// Tests for MONETcommon.FB_MonetTempSensor, the scaling and wire-break check of the 0-10 V temperature sensors.
// Cabinet_Over_Temp_Requests_Roof_Close: the cabinet temperature thresholds of MONETcommon.FB_MonetCabinetControl (BT1, driven
// through FB_MonetCabinetProbe) and its bCloseRoofRequest (#24 D9); no telescope is passed, so nothing is parked.
// Cabinet_Reads_The_Key_And_Passes_The_Safety_Inputs: FB_MonetCabinetControl as BROTLib.I_Cabinet (X1).
// Safety_Items_Decode_The_Info_Blocks: FB_MonetSafetyHandling as BROTLib.I_SafetyDiagnostics (X4), driven through FB_MonetSafetyProbe.
FUNCTION_BLOCK FB_MonetTempSensor_Tests EXTENDS TcUnit.FB_TestSuite
VAR
	nullComm	: FB_NullComm;
END_VAR

Mid_Scale_Is_Valid();
Wire_Break_Is_Invalid();
Over_Range_Is_Invalid();
Recovers_After_Wire_Break();
Cabinet_Over_Temp_Requests_Roof_Close();
Cabinet_Reads_The_Key_And_Passes_The_Safety_Inputs();
Safety_Items_Decode_The_Info_Blocks();

// 16384 of 32767 is 5 V, i.e. 25 C.
METHOD PRIVATE Mid_Scale_Is_Valid
VAR
	sensor	: MONETcommon.FB_MonetTempSensor;
END_VAR
TEST('Mid_Scale_Is_Valid');
sensor(iRaw := 16384, sName := 'TEMP_M1', comm := nullComm);
AssertTrue(Condition := sensor.bValid, Message := 'valid');
AssertEquals_REAL(Expected := 25.0, Actual := sensor.fTemperature, Delta := 0.01, Message := 'temperature');
TEST_FINISHED();
END_METHOD

// A broken wire reads about 0 V, which scales to -50 C.
METHOD PRIVATE Wire_Break_Is_Invalid
VAR
	sensor	: MONETcommon.FB_MonetTempSensor;
END_VAR
TEST('Wire_Break_Is_Invalid');
sensor(iRaw := 0, sName := 'TEMP_M1', comm := nullComm);
AssertFalse(Condition := sensor.bValid, Message := 'raw 0');
sensor(iRaw := 327, sName := 'TEMP_M1', comm := nullComm);
AssertFalse(Condition := sensor.bValid, Message := 'raw 327, just below 1 %');
sensor(iRaw := 328, sName := 'TEMP_M1', comm := nullComm);
AssertTrue(Condition := sensor.bValid, Message := 'raw 328, 1 %');
TEST_FINISHED();
END_METHOD

METHOD PRIVATE Over_Range_Is_Invalid
VAR
	sensor	: MONETcommon.FB_MonetTempSensor;
END_VAR
TEST('Over_Range_Is_Invalid');
sensor(iRaw := 32766, sName := 'TEMP_M1', comm := nullComm);
AssertTrue(Condition := sensor.bValid, Message := 'raw 32766');
sensor(iRaw := 32767, sName := 'TEMP_M1', comm := nullComm);
AssertFalse(Condition := sensor.bValid, Message := 'raw 32767, full scale');
TEST_FINISHED();
END_METHOD

METHOD PRIVATE Recovers_After_Wire_Break
VAR
	sensor	: MONETcommon.FB_MonetTempSensor;
END_VAR
TEST('Recovers_After_Wire_Break');
sensor(iRaw := 0, sName := 'TEMP_M1', comm := nullComm);
AssertFalse(Condition := sensor.bValid, Message := 'broken');
sensor(iRaw := 16384, sName := 'TEMP_M1', comm := nullComm);
AssertTrue(Condition := sensor.bValid, Message := 'reconnected');
TEST_FINISHED();
END_METHOD

// #24 D9 (owner decision: a critical cabinet temperature parks everything, the roof included): bCloseRoofRequest equals
// bCabinetOverTemp, set above 60 C and held until below 50 C, not latched beyond that. One call per temperature (BT1 in
// 0.1 C), no telescope (iTelescope 0).
METHOD PRIVATE Cabinet_Over_Temp_Requests_Roof_Close
VAR
	fbComm	: FB_NullComm;
	fbCab	: FB_MonetCabinetProbe(comm := fbComm);
END_VAR
TEST('Cabinet_Over_Temp_Requests_Roof_Close');
fbCab(fCabinetTempIn := 25.0);
AssertFalse(Condition := fbCab.bCloseRoofRequest, Message := '25 C: no roof close request');
fbCab(fCabinetTempIn := 59.9);
AssertFalse(Condition := fbCab.bCloseRoofRequest, Message := '59.9 C on the way up: no roof close request');
AssertFalse(Condition := fbCab.bCabinetOverTemp, Message := '59.9 C on the way up: not over temperature');
fbCab(fCabinetTempIn := 60.1);
AssertTrue(Condition := fbCab.bCloseRoofRequest, Message := '60.1 C: roof close requested');
AssertTrue(Condition := fbCab.bCabinetOverTemp, Message := '60.1 C: over temperature');
fbCab(fCabinetTempIn := 55.0);
AssertTrue(Condition := fbCab.bCloseRoofRequest, Message := '55 C on the way down: the request holds');
fbCab(fCabinetTempIn := 50.0);
AssertTrue(Condition := fbCab.bCloseRoofRequest, Message := '50.0 C on the way down: the request holds (reset below 50)');
fbCab(fCabinetTempIn := 49.9);
AssertFalse(Condition := fbCab.bCloseRoofRequest, Message := '49.9 C: the request is gone');
AssertFalse(Condition := fbCab.bCabinetOverTemp, Message := '49.9 C: not over temperature');
fbCab(fCabinetTempIn := 55.0);
AssertFalse(Condition := fbCab.bCloseRoofRequest, Message := '55 C on the way up again: no latch, no request');
TEST_FINISHED();
END_METHOD

// X1: ControlMode follows the Local/Remote key (inKeyLocal TRUE = Local), SwitchPresent is TRUE, the four other properties are the inputs.
METHOD PRIVATE Cabinet_Reads_The_Key_And_Passes_The_Safety_Inputs
VAR
	fbComm	: FB_NullComm;
	fbCab	: FB_MonetCabinetProbe(comm := fbComm);
	ipCab	: BROTLib.I_Cabinet;
END_VAR
TEST('Cabinet_Reads_The_Key_And_Passes_The_Safety_Inputs');
ipCab := fbCab;
fbCab(fCabinetTempIn := 25.0, bKeyLocalIn := FALSE, bEstop := FALSE, bSafetyError := FALSE, bSafetyAckPending := FALSE, bPendantActive := FALSE);
AssertTrue(Condition := ipCab.ControlMode = BROTLib.E_ControlMode.remote, Message := 'key off: Remote');
AssertTrue(Condition := ipCab.SwitchPresent, Message := 'the key is a physical switch');
AssertFalse(Condition := ipCab.EstopActive OR ipCab.SafetyError OR ipCab.SafetyAckPending OR ipCab.PendantActive, Message := 'inputs at rest: all FALSE');
fbCab(fCabinetTempIn := 25.0, bKeyLocalIn := TRUE, bEstop := FALSE, bSafetyError := FALSE, bSafetyAckPending := FALSE, bPendantActive := FALSE);
AssertTrue(Condition := ipCab.ControlMode = BROTLib.E_ControlMode.local, Message := 'key on: Local');
fbCab(fCabinetTempIn := 25.0, bKeyLocalIn := FALSE, bEstop := TRUE, bSafetyError := FALSE, bSafetyAckPending := FALSE, bPendantActive := FALSE);
AssertTrue(Condition := ipCab.EstopActive AND NOT ipCab.SafetyError AND NOT ipCab.SafetyAckPending AND NOT ipCab.PendantActive, Message := 'only EstopActive');
fbCab(fCabinetTempIn := 25.0, bKeyLocalIn := FALSE, bEstop := FALSE, bSafetyError := TRUE, bSafetyAckPending := FALSE, bPendantActive := FALSE);
AssertTrue(Condition := ipCab.SafetyError AND NOT ipCab.EstopActive AND NOT ipCab.SafetyAckPending AND NOT ipCab.PendantActive, Message := 'only SafetyError');
fbCab(fCabinetTempIn := 25.0, bKeyLocalIn := FALSE, bEstop := FALSE, bSafetyError := FALSE, bSafetyAckPending := TRUE, bPendantActive := FALSE);
AssertTrue(Condition := ipCab.SafetyAckPending AND NOT ipCab.EstopActive AND NOT ipCab.SafetyError AND NOT ipCab.PendantActive, Message := 'only SafetyAckPending');
fbCab(fCabinetTempIn := 25.0, bKeyLocalIn := FALSE, bEstop := FALSE, bSafetyError := FALSE, bSafetyAckPending := FALSE, bPendantActive := TRUE);
AssertTrue(Condition := ipCab.PendantActive AND NOT ipCab.EstopActive AND NOT ipCab.SafetyError AND NOT ipCab.SafetyAckPending, Message := 'only PendantActive');
TEST_FINISHED();
END_METHOD

// X4: items, texts, raw bytes, bOk, RestartPending (state RESET) and the derived StoActive, through the info data of the TwinSAFE blocks.
METHOD PRIVATE Safety_Items_Decode_The_Info_Blocks
VAR
	fbComm	: FB_NullComm;
	fbSafe	: FB_MonetSafetyProbe(comm := fbComm);
	ipSafe	: BROTLib.I_SafetyDiagnostics;
	stItems	: BROTLib.ST_SafetyItems;
END_VAR
TEST('Safety_Items_Decode_The_Info_Blocks');
ipSafe := fbSafe;
// everything in its normal running state
fbSafe(nGroupState := 1, nEStopState := 1, nEStopDiag := 0, nInState := 104, nInDiag := 0, nInSignals := 0, nOutState := 104, nOutDiag := 0, nOutSignals := 0);
stItems := ipSafe.Items;
AssertTrue(Condition := stItems.nCount = 4, Message := 'four items');
AssertEquals_STRING(Expected := 'safety.group1', Actual := stItems.aItem[1].sName, Message := 'item 1 name');
AssertEquals_STRING(Expected := 'safety.estop1', Actual := stItems.aItem[2].sName, Message := 'item 2 name');
AssertEquals_STRING(Expected := 'safety.el1904', Actual := stItems.aItem[3].sName, Message := 'item 3 name');
AssertEquals_STRING(Expected := 'safety.el2904', Actual := stItems.aItem[4].sName, Message := 'item 4 name');
AssertTrue(Condition := stItems.aItem[1].eKind = BROTLib.E_SafetyItemKind.group AND stItems.aItem[2].eKind = BROTLib.E_SafetyItemKind.estop
	AND stItems.aItem[3].eKind = BROTLib.E_SafetyItemKind.connection_in AND stItems.aItem[4].eKind = BROTLib.E_SafetyItemKind.connection_out, Message := 'kinds');
AssertTrue(Condition := stItems.aItem[1].bOk AND stItems.aItem[2].bOk AND stItems.aItem[3].bOk AND stItems.aItem[4].bOk, Message := 'all ok in the normal state');
AssertEquals_STRING(Expected := 'RUN', Actual := stItems.aItem[1].sState, Message := 'group state text');
AssertEquals_STRING(Expected := 'State Data', Actual := stItems.aItem[3].sState, Message := 'connection state text');
AssertFalse(Condition := ipSafe.StoActive, Message := 'no STO in the normal state');
AssertFalse(Condition := ipSafe.RestartPending, Message := 'no restart pending in the normal state');
// E-stop pressed: state STOP
fbSafe(nGroupState := 1, nEStopState := 2, nEStopDiag := 0, nInState := 104, nInDiag := 0, nInSignals := 0, nOutState := 104, nOutDiag := 0, nOutSignals := 0);
stItems := ipSafe.Items;
AssertFalse(Condition := stItems.aItem[2].bOk, Message := 'E-stop item not ok');
AssertEquals_STRING(Expected := 'STOP', Actual := stItems.aItem[2].sState, Message := 'E-stop state text');
AssertTrue(Condition := stItems.aItem[2].nMapState = 2, Message := 'raw E-stop map state');
AssertTrue(Condition := stItems.aItem[1].bOk, Message := 'the group item is not affected');
AssertTrue(Condition := ipSafe.StoActive, Message := 'STO derived from the E-stop not in RUN');
AssertFalse(Condition := ipSafe.RestartPending, Message := 'STOP is not RESET');
// group waits for restart: state RESET (also with the E-stop function)
fbSafe(nGroupState := 5, nEStopState := 5, nEStopDiag := 0, nInState := 104, nInDiag := 0, nInSignals := 0, nOutState := 104, nOutDiag := 0, nOutSignals := 0);
stItems := ipSafe.Items;
AssertTrue(Condition := ipSafe.RestartPending, Message := 'RESET: restart pending');
AssertEquals_STRING(Expected := 'RESET', Actual := stItems.aItem[1].sState, Message := 'group state text RESET');
AssertFalse(Condition := stItems.aItem[1].bOk, Message := 'group item not ok in RESET');
AssertTrue(Condition := ipSafe.StoActive, Message := 'STO derived');
// only the E-stop function waits
fbSafe(nGroupState := 1, nEStopState := 5, nEStopDiag := 0, nInState := 104, nInDiag := 0, nInSignals := 0, nOutState := 104, nOutDiag := 0, nOutSignals := 0);
AssertTrue(Condition := ipSafe.RestartPending, Message := 'E-stop RESET alone: restart pending');
// a diagnosis on the E-stop makes it not ok even in RUN
fbSafe(nGroupState := 1, nEStopState := 1, nEStopDiag := 16, nInState := 104, nInDiag := 0, nInSignals := 0, nOutState := 104, nOutDiag := 0, nOutSignals := 0);
stItems := ipSafe.Items;
AssertFalse(Condition := stItems.aItem[2].bOk, Message := 'E-stop diagnosis: not ok');
AssertEquals_STRING(Expected := 'EDM Error EDM 1', Actual := stItems.aItem[2].sDiag, Message := 'E-stop diagnosis text');
// connections: diagnosis, channel bits (low nibble only), other state
fbSafe(nGroupState := 1, nEStopState := 1, nEStopDiag := 0, nInState := 104, nInDiag := 5, nInSignals := 245, nOutState := 103, nOutDiag := 0, nOutSignals := 0);
stItems := ipSafe.Items;
AssertFalse(Condition := stItems.aItem[3].bOk, Message := 'EL1904 diagnosis: not ok');
AssertEquals_STRING(Expected := 'Watchdog expired', Actual := stItems.aItem[3].sDiag, Message := 'EL1904 diagnosis text');
AssertTrue(Condition := stItems.aItem[3].nChannels = 16#05, Message := 'EL1904 channels 1 and 3');
AssertTrue(Condition := stItems.aItem[3].nMapDiag = 16#05, Message := 'raw EL1904 diagnosis');
AssertFalse(Condition := stItems.aItem[4].bOk, Message := 'EL2904 not in State Data');
AssertEquals_STRING(Expected := 'State Parameter', Actual := stItems.aItem[4].sState, Message := 'EL2904 state text');
TEST_FINISHED();
END_METHOD

END_FUNCTION_BLOCK

(* stored: Version 1.1.0.1, ProductVersion 3.1.4024.15
   POU FB_MonetTempSensor_Tests: Id {2c9e5b17-f4a8-4d03-b6e1-93a07d58c2f4}, SpecialFunc None
   Method Mid_Scale_Is_Valid: Id {a4d17c3e-8b25-4f60-91ce-5e2b7a0d3c18}
   Method Wire_Break_Is_Invalid: Id {e61b08f9-37d4-4a52-8c7a-1d9f40b6e253}
   Method Over_Range_Is_Invalid: Id {57f2c9a0-1e6b-4d38-a3b7-c08d9e41f762}
   Method Recovers_After_Wire_Break: Id {b83e6d15-9c40-4a7f-82d1-f5a60c2e9b37}
   Method Cabinet_Over_Temp_Requests_Roof_Close: Id {3f4047b1-637c-49e1-aad4-048bd6bd5304}
   Method Cabinet_Reads_The_Key_And_Passes_The_Safety_Inputs: Id {eab4d8e2-9d21-4636-93cc-4a6fe8561573}
   Method Safety_Items_Decode_The_Info_Blocks: Id {ede2ebd7-8118-4e99-91f3-597f21ae7353} *)
